# EPICS autosave request: 1.5.0/debian-12/7.0.10/modules/ADCore-ee039d2/db/ADAutoSaveMenu.req
file "configMenu_settings.req", P=$(P), CONFIG=ADAutoSave
file "auto_settings.req", P=$(P)
